Staubli VAL3: main.pgx

program main()
begin
  close(tCurrentTool)
  pPointRx.config.shoulder = lefty
  pPointRx.config.elbow = epositive
  pPointRx.config.wrist = wpositive
  pPointRx2.config.shoulder = lefty
  pPointRx2.config.elbow = epositive
  pPointRx2.config.wrist = wpositive
  mCurrentSpeed.tvel = 100.00
  mCurrentSpeed.blend = joint
  mCurrentSpeed.reach = 0.010
  mCurrentSpeed.leave = 0.010
  // Program SplitTest start
  // Program generated by VerticalBot Studio for Staubli RX160 on 25/10/2026 12:00:00
  // Using nominal kinematics.
  mCurrentSpeed.tvel = 200.000
  call MoveJoint(10.00000,20.00000,90.00000,30.00000,45.00000,60.00000)
  call MoveLine(1077.300,-56.172,837.243,-146.156,25.288,-102.118)
  call MoveLine(1005.190,-118.362,847.372,-147.806,26.655,-97.799)
  call MoveLine(1077.300,-56.172,837.243,-146.156,25.288,-102.118)
  call MoveLine(1005.190,-118.362,847.372,-147.806,26.655,-97.799)
  call MoveLine(1077.300,-56.172,837.243,-146.156,25.288,-102.118)
  call MoveLine(1005.190,-118.362,847.372,-147.806,26.655,-97.799)
  call MoveLine(1077.300,-56.172,837.243,-146.156,25.288,-102.118)
  call MoveLine(1005.190,-118.362,847.372,-147.806,26.655,-97.799)
  call MoveLine(1077.300,-56.172,837.243,-146.156,25.288,-102.118)
  call MoveLine(1005.190,-118.362,847.372,-147.806,26.655,-97.799)

end
